// TIA Portal V17 export
FUNCTION_BLOCK "FB_T04c_CTU"   // FB143, LAD
{ S7_Optimized_Access := 'TRUE' }
// stored: IsIECCheckEnabled false, MemoryReserve 100, SetENOAutomatically false
   VAR_INPUT
      Impulsion : Bool;
      RAZ : Bool;
      Consigne : Int;
   END_VAR
   VAR_OUTPUT
      Atteint : Bool;
      Compte : Int;
   END_VAR
   VAR
      ctuPieces : CTU_INT;
   END_VAR
BEGIN

REGION Network 1: Compteur CTU
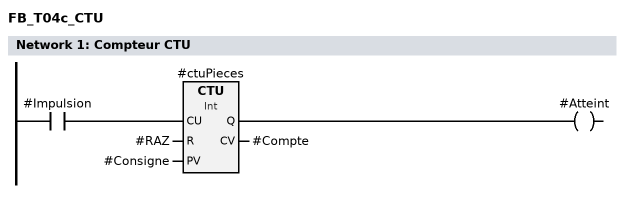
   RUNG wire#powerrail
      Contact( #Impulsion )
      { S7_Templates := "value_type := Int" } #ctuPieces.CTU(r := #RAZ, pv := #Consigne, cv => #Compte)
      Coil( #Atteint )
   END_RUNG
   // the same network as SCL:
   #ctuPieces(CU := #Impulsion, R := #RAZ, PV := #Consigne, CV => #Compte);   // CTU
   #Atteint := #ctuPieces.Q;
END_REGION
END_FUNCTION_BLOCK
